(* PLC project EnhancedSystemWithCounter, PLCArchitect Machine Expert Logic Builder V19.2.3.0 *)
(* stored: creationDateTime 2026-02-05T20:35:55.192173, version 1.0.0.0 *)

PROGRAM EnhancedSystemWithCounter
  VAR
    StartBtn : BOOL;
    ProcessActive : BOOL;
    AgitatorMotor : BOOL;
    HeatingElement : BOOL;
    MixingTimer : TON;
    HeatingTimer : TON;
    MixingTime : TIME;
    HeatingTime : TIME;
    BatchCounter : CTU;
    CounterReset : BOOL;
    BatchTarget : INT;
    BatchComplete : BOOL;
    TempController : PID_FIXCYCLE;
    actual_temp : REAL;
    setpoint_temp : REAL;
    Manual : BOOL;
    reset : BOOL;
    y_manual : REAL;
    y_offset : REAL;
    y_min : REAL;
    y_max : REAL;
    cycle : REAL;
    limits_active : BOOL;
    Overflow : BOOL;
    heater_output : REAL;
  END_VAR
  VAR  (* added by the conversion: wires and edge detectors of the diagram *)
    F_TRIG1 : F_TRIG;
  END_VAR

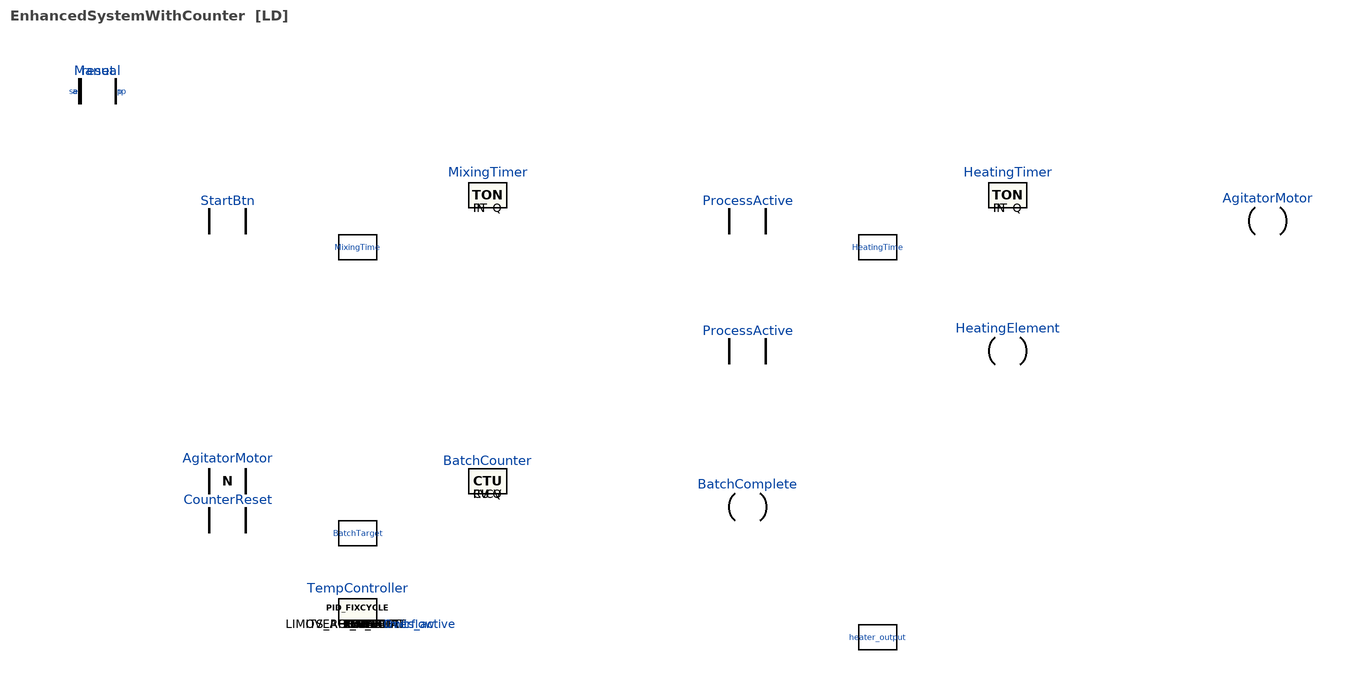
(* LD diagram, written out as Structured Text *)
MixingTimer(IN := StartBtn, PT := MixingTime);
HeatingTimer(IN := MixingTimer.Q AND ProcessActive, PT := HeatingTime);
AgitatorMotor := HeatingTimer.Q;
HeatingElement := ProcessActive;
F_TRIG1(CLK := AgitatorMotor);
BatchCounter(CU := F_TRIG1.Q, R := CounterReset, PV := BatchTarget);
BatchComplete := BatchCounter.Q;
TempController(ACTUAL := actual_temp, SET_POINT := setpoint_temp, KP := 1.5, TN := 10.0, TV := 2.0, Y_MANUAL := y_manual, Y_OFFSET := y_offset, Y_MIN := y_min, Y_MAX := y_max, MANUAL := Manual, RESET := reset, CYCLE := cycle, LIMITS_ACTIVE => limits_active, OVERFLOW => Overflow);
heater_output := TempController.Y;
END_PROGRAM
